Fanuc KAREL source: kb00133.KL

-- PROVISIONAL review KL for V770-1; original PC SHA256 4885083bfe34e8f877aa93c4a874b682f76320ad7a5209d47a5386be17bc1476
-- Incomplete behavior may be omitted. Consult companion uncertainty JSON. Do not deploy.
PROGRAM KB00133
%NOLOCKGROUP
BEGIN
  -- UNRESOLVED_PC offsets 5-12; opcodes 9D,23
  -- UNRESOLVED_PC offsets 17-24; opcodes 9D,23
  -- UNRESOLVED_PC offsets 29-36; opcodes 9D,23
  -- UNRESOLVED_PC offsets 41-48; opcodes 9D,23
  -- UNRESOLVED_PC offsets 53-60; opcodes 9D,23
  -- UNRESOLVED_PC offsets 65-99; opcodes 27,22,22,22,22,22,31
  -- UNRESOLVED_PC offsets 104-108; opcodes 7F
END KB00133
